(* IEC 61131-3 sources: llm-plc-st-eval/data/processed_definitivo/claude-sonnet-4-6/B7/few_shot, 3 files *)

(* ---- ejec_1.st ---- *)
FUNCTION SelBomba : BOOL
VAR_INPUT
    modoAuto  : BOOL; (* TRUE = modo automatico, FALSE = modo manual *)
    btnManual : BOOL; (* Boton de mando manual de la bomba *)
    nivelBajo : BOOL; (* Senal de nivel bajo del deposito *)
END_VAR

(* Sin memoria entre ciclos: el resultado depende solo de las entradas actuales *)
(* En modo automatico la bomba sigue a nivelBajo; en manual sigue a btnManual *)
SelBomba := (modoAuto AND nivelBajo) OR (NOT modoAuto AND btnManual);
END_FUNCTION

(* ---- ejec_2.st ---- *)
FUNCTION SelBomba : BOOL
VAR_INPUT
    modoAuto  : BOOL; (* TRUE = modo automatico, FALSE = modo manual *)
    btnManual : BOOL; (* Boton de mando en modo manual *)
    nivelBajo : BOOL; (* Senal de nivel bajo del deposito *)
END_VAR

(* Sin memoria entre ciclos: el resultado depende solo de las entradas actuales *)
(* En modo automatico la bomba sigue a nivelBajo; en manual sigue a btnManual *)
SelBomba := (modoAuto AND nivelBajo) OR (NOT modoAuto AND btnManual);
END_FUNCTION

(* ---- ejec_3.st ---- *)
FUNCTION SelBomba : BOOL
VAR_INPUT
    modoAuto  : BOOL; (* TRUE = modo automatico, FALSE = modo manual *)
    btnManual : BOOL; (* Boton de mando manual de la bomba *)
    nivelBajo : BOOL; (* Senal de nivel bajo del deposito *)
END_VAR

(* Sin memoria entre ciclos: el resultado depende solo de las entradas actuales *)
(* Modo automatico: bomba encendida si hay nivel bajo                          *)
(* Modo manual    : bomba obedece directamente al boton                        *)
SelBomba := (modoAuto AND nivelBajo) OR (NOT modoAuto AND btnManual);
END_FUNCTION
